FUNCTION_BLOCK MotorBaseNer_HMI (* Service Interface Function Block Type *)
  (* Standard: 61499-2 *)
  (* Version 1.0.1, 1/30/2024, ApplicationLibDevTeam, Schneider Electric, First Version *)
  PACKAGE SE.Nereda;
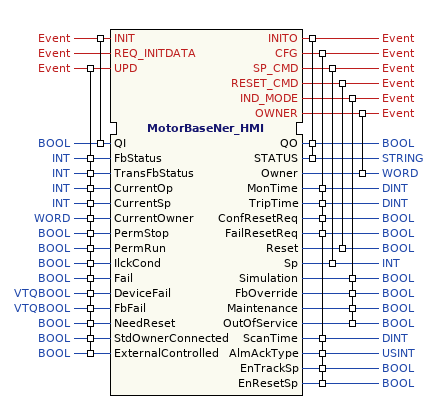
  EVENT_INPUT
    INIT WITH QI;
    REQ_INITDATA; (* Request to initialize data *)
    UPD WITH FbStatus, TransFbStatus, CurrentOp, CurrentSp, NeedReset, FbFail, DeviceFail, IlckCond, PermStop, PermRun, Fail, CurrentOwner, StdOwnerConnected, ExternalControlled; (* Update data to supervision *)
  END_EVENT
  EVENT_OUTPUT
    INITO WITH QO, STATUS;
    CFG WITH MonTime, TripTime, ConfResetReq, FailResetReq, ScanTime, AlmAckType, EnTrackSp, EnResetSp; (* Request for new parameter *)
    SP_CMD WITH Sp; (* Request for new operator setpoint *)
    RESET_CMD WITH Reset; (* Request to reset device *)
    IND_MODE WITH Simulation, FbOverride, Maintenance, OutOfService; (* Request for new operational modes *)
    OWNER WITH Owner; (* Request for owner change *)
  END_EVENT
  VAR_INPUT
    QI : BOOL;
    FbStatus : INT; (* Device state(0 = stopped, 1= Running) *) {SET_ATTRIBUTE(Runtime.Archive.Counters, AbsoluteValues=False)} {SET_ATTRIBUTE(Runtime.Archive.Id, 1)} {SET_ATTRIBUTE(Runtime.History.Depth, 100)} {SET_ATTRIBUTE(Runtime.History.SmoothTime, 60000)} {SET_ATTRIBUTE(Runtime.History.SmoothValue, 1)}
    TransFbStatus : INT; (* Device transition state( 0 = Stopped, 1 = Running, 5 = Stopping , 6 = Starting and 253 = Unknown) *) {SET_ATTRIBUTE(Runtime.Archive.Counters, AbsoluteValues=False)} {SET_ATTRIBUTE(Runtime.Archive.Id, 1)} {SET_ATTRIBUTE(Runtime.History.Depth, 100)} {SET_ATTRIBUTE(Runtime.History.SmoothTime, 60000)} {SET_ATTRIBUTE(Runtime.History.SmoothValue, 1)}
    CurrentOp : INT; (* Current value of the output ( 0 = Stop command and 1 = start command) *) {SET_ATTRIBUTE(Runtime.Archive.Counters, AbsoluteValues=False)} {SET_ATTRIBUTE(Runtime.Archive.Id, 1)} {SET_ATTRIBUTE(Runtime.History.Depth, 100)} {SET_ATTRIBUTE(Runtime.History.SmoothTime, 60000)} {SET_ATTRIBUTE(Runtime.History.SmoothValue, 1)}
    CurrentSp : INT; (* Current value of the setpoint ( 0 = Stop Setpoint and 1 = start setpoint *) {SET_ATTRIBUTE(Runtime.Archive.Counters, AbsoluteValues=False)} {SET_ATTRIBUTE(Runtime.Archive.Id, 1)} {SET_ATTRIBUTE(Runtime.History.Depth, 100)} {SET_ATTRIBUTE(Runtime.History.SmoothTime, 60000)} {SET_ATTRIBUTE(Runtime.History.SmoothValue, 1)}
    CurrentOwner : WORD; (* Current Owner status ( 16#08 = Program remote  and 16#10 = Operator) *)
    PermStop : BOOL; (* 1= Stop permission available *)
    PermRun : BOOL; (* 1= Start permission available *)
    IlckCond : BOOL; (* 1= Interlock active *)
    Fail : BOOL; (* 1= Fail active *)
    DeviceFail : VTQBOOL; (* 1=Device fail alarm status active *)
    FbFail : VTQBOOL; (* 1=Feedback fail alarm status active *)
    NeedReset : BOOL; (* 1= Device need reset *)
    StdOwnerConnected : BOOL; (* 1= External owner connected *)
    ExternalControlled : BOOL; (* 1 = Device is externally controlled *)
  END_VAR
  VAR_OUTPUT
    QO : BOOL; (* Event Output Qualifier *)
    STATUS : STRING; (* Service Status *)
    Owner : WORD; (* Requested owner (16#10 = Operator, 16#8 = Program remote) *)
    MonTime : DINT; (* Feedback monitoring time *)
    TripTime : DINT; (* Feedback trip time *)
    ConfResetReq : BOOL; (* 1= Need reset on confirmation mismatch *)
    FailResetReq : BOOL; (* 1 = Need reset on device detected failure *)
    Reset : BOOL; (* 1 = Reset request from supervision *)
    Sp : INT; (* New setpoint from the supervision *)
    Simulation : BOOL; (* 1 = Enable device in simulation *)
    FbOverride : BOOL; (* 1 = Enable device in override mode *)
    Maintenance : BOOL; (* 1 = Enable device in maintenance mode *)
    OutOfService : BOOL; (* 1 = Enable device in out of service mode *)
    ScanTime : DINT; (* Alarm holding time *)
    AlmAckType : USINT; (* 0=Not ackable; 1=Ack deletes; 2=Came has to be acked; 3=Came and gone have to be acked; 4=Pair has to be acked *)
    EnTrackSp : BOOL; (* 1= Enable the tracking of Interlock setpoint *)
    EnResetSp : BOOL; (* 1= Enable Reset Setpoint *)
  END_VAR
  SERVICE /
    SEQUENCE 
    END_SEQUENCE
  END_SERVICE
END_FUNCTION_BLOCK
